// TIA Portal V19 export
TYPE "ST_SAF"
   STRUCT
      EMG : "ST_EMG";
      FENCE : "ST_FENCE";
      DOOR : "ST_DOOR";
      ZONE : "ST_SAFETY_ZONE";
   END_STRUCT;
END_TYPE
